Fanuc KAREL source: KB00052.KL

PROGRAM KB00052
%NOLOCKGROUP
VAR
  P1: INTEGER
  P2: INTEGER
  RESULT: XYZWPREXT
BEGIN
  P1 = 1
  P2 = 1
  RESULT = CURPOS(P1, P2)
END KB00052
